Fanuc KAREL source: KB00167.KL

PROGRAM KB00167
%NOLOCKGROUP
VAR
  P1: INTEGER
  P2: INTEGER
  P3: JOINTPOS
  P4: INTEGER
BEGIN
  P1 = 1
  P2 = 1
  P4 = 1
  SET_JPOS_TPE(P1, P2, P3, P4)
END KB00167
